Fanuc KAREL source: kb00037.KL

-- PROVISIONAL review KL for V940-1; original PC SHA256 f90cfc98d1836946eff56f41262e3533de708df3e4a097042feee9cd28d05e33
-- Incomplete behavior may be omitted. Consult companion uncertainty JSON. Do not deploy.
PROGRAM KB00037
%NOLOCKGROUP
BEGIN
  -- V9_ZERO_TABLE_METADATA_HINT layout=0002_ascii; no indexed target words; source/name/runtime held
  -- UNRESOLVED_PC offsets 5-16; opcodes 2E,23
  -- UNRESOLVED_PC offsets 21-28; opcodes 9D,23
  -- UNRESOLVED_PC offsets 33-40; opcodes 9D,23
  -- UNRESOLVED_PC offsets 45-54; opcodes 3F,75
  -- UNRESOLVED_PC offsets 59-89; opcodes 27,22,22,22,22,2A,31
  -- UNRESOLVED_PC offsets 94-98; opcodes 7F
END KB00037
